(* IEC 61131-3 sources: Caravan/Archiv/12-04-19/Stations/MachineControl/MachineControl/Class/AmpFilter_Class, 1 file *)

(* ---- AmpFilter_Class.st ---- *)
(*!
<Class
	Name               = "AmpFilter_Class"
	Revision           = "0.0"
	RealtimeTask       = "true"
	CyclicTask         = "false"
	BackgroundTask     = "false"
	Sigmatek           = "false"
	OSInterface        = "false"
	HighPriority       = "false"
	Automatic          = "false"
	UpdateMode         = "Prescan"
	SharedCommandTable = "true"
	Objectsize         = "(570,180)">
	<Channels>
		<Server Name="ClassSvr" Visualized="false" Initialize="false" WriteProtected="true" Retentive="false"/>
		<Server Name="CorrectedOutput_S" Visualized="false" Initialize="false" WriteProtected="true" Retentive="false"/>
		<Client Name="VoltageImput1_C" Required="true" Internal="false"/>
		<Client Name="VoltageImput2_C" Required="true" Internal="false"/>
	</Channels>
</Class>
*)
AmpFilter_Class : CLASS
	TYPE
	  Type0 : ARRAY [0..999] OF DINT;
	END_TYPE
  //Servers:
	ClassSvr 	: SvrChCmd_DINT;
	CorrectedOutput_S 	: SvrCh_DINT;
  //Clients:
	VoltageImput1_C 	: CltCh_DINT;
	VoltageImput2_C 	: CltCh_DINT;
  //Variables:
		Counter_VAR 	: DINT;
		DataArray : ARRAY [0..999] OF DINT;

  //Functions:

	FUNCTION VIRTUAL GLOBAL RtWork
		VAR_INPUT
			EAX 	: UDINT;
		END_VAR
		VAR_OUTPUT
			state (EAX) 	: UDINT;
		END_VAR;
  //Tables:
	FUNCTION @STD
		VAR_OUTPUT
			ret_code	: CONFSTATES;
		END_VAR;
	FUNCTION GLOBAL TAB @CT_;
END_CLASS;

FUNCTION VIRTUAL GLOBAL AmpFilter_Class::RtWork
	VAR_INPUT
		EAX 	: UDINT;
	END_VAR
	VAR_OUTPUT
		state (EAX) 	: UDINT;
	END_VAR

  //Read in
  VoltageImput1_C   :=  VoltageImput1_C.Read();
  VoltageImput2_C   :=  VoltageImput2_C.Read();

  for Counter_VAR := 0 to 999 by 1 do

      DataArray[Counter_VAR] :=  VoltageImput1_C;

  end_for;

	state := READY;

END_FUNCTION
